Yaskawa INFORM job: PGPROG.JBI

/JOB
//NAME PGPROG
//POS
///NPOS 11,0,0,0,0,0
///TOOL 9
///POSTYPE PULSE
///PULSE
C00000=0,-10240,0,-34475,0,0,22983
C00001=0,-10240,0,-34475,0,0,22983
C00002=0,-10240,0,-34475,0,0,22983
C00003=0,-10240,0,-34475,0,0,22983
C00004=0,-10240,0,-34475,0,0,22983
C00005=20480,-10240,0,-34475,0,-8704,22983
C00006=0,-10240,0,-34475,0,0,22983
C00007=0,-10240,0,-34475,0,0,22983
C00008=0,-10240,0,-34475,0,0,22983
C00009=10240,-5120,-5746,-40220,-5746,-2901,28729
C00010=-5120,-5120,-11492,-45966,11492,-14507,17237
//INST
<volatile>
///COMM Generated using RoboDK
///ATTR SC,RW
///GROUP1 RB1
NOP
'Program generated by RoboDK v
'6.0.7 for Yaskawa Motoman CSD
'A10F on XX/XX/XXXX 18:00:00
'Using nominal kinematics.
'Using Frame Pg (targets wrt b
'ase):
'1234.6,-98.8,50.5,0.0,0.0,30.
'0
'Tool Tool Pg should be close
'to:
'10.0,20.0,150.0,15.0,0.0,0.0
MOVJ C00000 VJ=50.00 PL=5
MOVL C00001 V=250.0 PL=5
MOVC C00002 V=250.0 PL=5
MOVC C00003 V=250.0 PL=5
MOVC C00004 V=250.0 PL=5
MOVJ C00005 VJ=50.00 PL=5
MOVL C00006 V=100.0 ACC=100 DEC=100
MOVL C00007 V=100.0 ACC=100 DEC=100
TIMER T=0.50
PAUSE
MSG "Hello from postgen"
'a comment
CALL JOB:SUBPROG
CustomCode(42)
ThreadProg
DOUT OT#(1) ON
DOUT Valve OFF
DOUT OT#(3) 2.5
WAIT IN#(2)=ON
WAIT IN#(4)=OFF T=1.50
'Tool Tool2 should be close to
':
'0.0,0.0,200.0,0.0,0.0,0.0
MOVJ C00008 VJ=60.00 ACC=100 DEC=100
MOVJ C00009 VJ=60.00 ACC=100 DEC=100
MOVL C00010 V=100.0 ACC=100 DEC=100
END
